FUNCTION_BLOCK b_abs
VAR_INPUT
	x: ARRAY[0..2] OF LREAL;
END_VAR
VAR_OUTPUT
	y: ARRAY[0..2] OF LREAL;
END_VAR
VAR
END_VAR


y[0] := ABS(x[0]);
y[1] := ABS(x[1]);
y[2] := ABS(x[2]);

END_FUNCTION_BLOCK

(* stored: Version 1.1.0.1, ProductVersion 3.1.4024.9
   POU b_abs: Id {0159dded-4d7f-4927-9919-ac36ca379040}, SpecialFunc None *)
